// TIA Portal V15.1 export
// export: Created 2026-11-01T20:56:25.3861065Z, ExportSetting WithDefaults, DisplayName Totally Integrated Automation Portal, DisplayVersion V15.1, DisplayName TIA Portal Openness, DisplayVersion V15.1, DisplayName STEP 7 Professional, DisplayVersion V15.1, DisplayName WinCC Professional, DisplayVersion V15.1
TagTable "Default tag table"
  Par_SP : Int  (PLC tag Par.SP, HMI_Connection_1, 1 s)
